(* IEC 61131-3 sources: trust-platform/examples/OSCAT/solar_lighting_clock/non-oop/src, 1 file *)

(* ---- Configuration.st ---- *)
CONFIGURATION SolarLightingClockClassicConfiguration
RESOURCE SolarLightingClockClassic ON PLC
    TASK MainTask (INTERVAL := T#1s, PRIORITY := 1);
    PROGRAM Main WITH MainTask : Main;
END_RESOURCE
END_CONFIGURATION
